(* IEC 61131-3 sources: Zbiorniki_user/Temp/Import/MpFile, 4 files *)

(* ---- MpFile.typ ---- *)
TYPE
	MpFileManagerUIItemType : 	STRUCT
		Name : STRING[255]; (*Filename / Folder name*)
		Size : UDINT; (*File size [bytes]*)
		LastModified : DATE_AND_TIME; (*Date when this file/folder was last modified*)
		ItemType : MpFileManagerUIItemTypeEnum; (*File type (.csv, .jpg, etc.)*)
		IsSelected : BOOL; (*Indicates that a file/folder is selected*)
		IsFolder : BOOL; (*Indicates that the element is a folder*)
	END_STRUCT;
	MpFileManagerUIItemTypeEnum :
		(
		mpFILE_ITEM_TYPE_NONE := 0, (*No type defined*)
		mpFILE_ITEM_TYPE_FOLDER := 1, (*Indicates that the element is a folder*)
		mpFILE_ITEM_TYPE_FILE := 2, (*Indicates that the element is a file*)
		mpFILE_ITEM_TYPE_TXT := 3, (*Indicates that the element is a text file*)
		mpFILE_ITEM_TYPE_HTML := 4, (*Indicates that the element is an HTML file*)
		mpFILE_ITEM_TYPE_DOC := 5, (*Indicates that the element is a Word file (.doc) *)
		mpFILE_ITEM_TYPE_XLS := 6, (*Indicates that the element is an Excel file (.xls)*)
		mpFILE_ITEM_TYPE_XML := 7, (*Indicates that the element is an XML file (.xml)*)
		mpFILE_ITEM_TYPE_CSV := 8, (*Indicates that the element is an CSV file (.csv)*)
		mpFILE_ITEM_TYPE_JPG := 9, (*Indicates that the element is an image file (.jpg)*)
		mpFILE_ITEM_TYPE_BMP := 10, (*Indicates that the element is an image file (.bmp)*)
		mpFILE_ITEM_TYPE_USER1 := 89, (*Indicates that the element is an user predefined type 1*)
		mpFILE_ITEM_TYPE_USER2 := 90, (*Indicates that the element is an user predefined type 2*)
		mpFILE_ITEM_TYPE_USER3 := 91, (*Indicates that the element is an user predefined type 3*)
		mpFILE_ITEM_TYPE_USER4 := 92, (*Indicates that the element is an user predefined type 4*)
		mpFILE_ITEM_TYPE_USER5 := 93, (*Indicates that the element is an user predefined type 5*)
		mpFILE_ITEM_TYPE_USER6 := 94, (*Indicates that the element is an user predefined type 6*)
		mpFILE_ITEM_TYPE_USER7 := 95, (*Indicates that the element is an user predefined type 7*)
		mpFILE_ITEM_TYPE_USER8 := 96, (*Indicates that the element is an user predefined type 8*)
		mpFILE_ITEM_TYPE_USER9 := 97, (*Indicates that the element is an user predefined type 9*)
		mpFILE_ITEM_TYPE_USER10 := 98, (*Indicates that the element is an user predefined type 10*)
		mpFILE_ITEM_TYPE_UNKNOWN := 99 (*Indicates that the file type is unknown*)
		);
	MpFileManagerUISortOrderEnum :
		(
		mpFILE_SORT_BY_NAME_ASC := 0, (*Sorts in ascending (alphabetic) order*)
		mpFILE_SORT_BY_NAME_DESC := 1, (*Sorts in descending (alphabetic) order*)
		mpFILE_SORT_BY_SIZE_ASC := 2, (*Sorts in ascending order by file size*)
		mpFILE_SORT_BY_SIZE_DES := 3, (*Sorts in descending order by file size*)
		mpFILE_SORT_BY_MOD_TIME_ASC := 4, (*Sorts in ascending order by date last modified*)
		mpFILE_SORT_BY_MOD_TIME_DESC := 5 (*Sorts in descending order by date last modified*)
		);
	MpFileManagerUIMessageEnum :
		(
		mpFILE_MSG_OK := 0, (*Dialog box for requesting confirmation of input*)
		mpFILE_MSG_CONFIRM_DELETE := 1, (*Dialog box for requesting confirmation of deletion*)
		mpFILE_MSG_CONFIRM_OVERWRITE := 2, (*Dialog box for requesting confirmation of overwriting*)
		mpFILE_MSG_BUSY := 3 (*Dialog box for requesting confirmation of busy UI*)
		);
	MpFileDiagType : 	STRUCT
		StatusID : MpFileStatusIDType; (*StatusID diagnostic structure*)
	END_STRUCT;
	MpFileStatusIDType : 	STRUCT
		ID : MpFileErrorEnum; (*Error code for mapp component*)
		Severity : MpComSeveritiesEnum; (*Describes the type of information supplied by the status ID (success, information, warning, error)*)
		Code : UINT; (*Code for the status ID. This error number can be used to search for additional information in the help system.*)
	END_STRUCT;
	MpFileInfoType : 	STRUCT
		Diag : MpFileDiagType; (*Diagnostic structure for the status ID*)
	END_STRUCT;
	MpFileManagerUIStatusEnum :
		(
		mpFILE_UI_STATUS_IDLE := 0, (*Indicates that no process is currently active*)
		mpFILE_UI_STATUS_REFRESH := 1, (*Updating elements*)
		mpFILE_UI_STATUS_CHANGE_PAGE := 2, (*Page change active*)
		mpFILE_UI_STATUS_CHANGE_DIR := 3, (*Folder change active*)
		mpFILE_UI_STATUS_CHANGE_DEVICE := 4, (*File Device Change active*)
		mpFILE_UI_STATUS_CREATE := 5, (*Creating a file/folder active*)
		mpFILE_UI_STATUS_RENAME := 6, (*Renaming a file/folder active*)
		mpFILE_UI_STATUS_DELETE := 7, (*Deleting a file/folder active*)
		mpFILE_UI_STATUS_COPY := 8, (*Copying a file/folder active*)
		mpFILE_UI_STATUS_CUT := 9, (*Cutting a file/folder active*)
		mpFILE_UI_STATUS_PASTE := 10, (*Pasting a file/folder active*)
		mpFILE_UI_STATUS_SORT := 11, (*Sorting files/folders in specified sort order*)
		mpFILE_UI_STATUS_ERROR := 99 (*The last operation generated an error*)
		);
	MpFileManagerUISetupType : 	STRUCT
		FileListSize : UINT := 10; (*Number of files to be displayed on one page of the list in the HMI application*)
		FileListScrollWindow : USINT := 1; (*Determines how many entries from the list are displayed in advance when scrolling up and down*)
	END_STRUCT;
	MpFileManagerUIConnectType : 	STRUCT
		Status : MpFileManagerUIStatusEnum; (*Current operation*)
		DeviceList : MpFileManagerUIDeviceListType; (*List of data storage media (file devices) accessible by the file manager*)
		File : MpFileManagerUIFileType; (*Contains the file list as well as additional information about files,folders and possible commands*)
		MessageBox : MpFileManagerUIMessageBoxType; (*Controls dialog boxes*)
		DefaultLayerStatus : UINT; (*Status DP for the default layer of the visu page where the file manager is being displayed*)
	END_STRUCT;
	MpFileManagerUIMessageBoxType : 	STRUCT
		LayerStatus : UINT; (*Visibility of the dialog box*)
		Type : MpFileManagerUIMessageEnum; (*Type of dialog box*)
		ErrorNumber : UINT; (*Current error number to be displayed*)
		Confirm : BOOL; (*Confirms the operation*)
		Cancel : BOOL; (*Cancels the operation*)
	END_STRUCT;
	MpFileManagerUIPathInfoType : 	STRUCT
		CurrentDir : STRING[255]; (*Current folder name*)
		FileCount : UDINT; (*Number of files in the current folder*)
		FolderCount : UDINT; (*Number of subfolders in the current folder*)
	END_STRUCT;
	MpFileManagerUIFileType : 	STRUCT
		List : MpFileManagerUIFileListType; (*List of all folders and files under the current path, as well as the navigation of the list*)
		Filter : STRING[255]; (*Filter used to sort the files*) (* *) (*#CMD#OPT#;*)
		SortOrder : MpFileManagerUISortOrderEnum; (*Responsible for the order of files in the list*)
		Refresh : BOOL; (*Updates the file list in the current folder*)
		PathInfo : MpFileManagerUIPathInfoType; (*Information about the current path*)
		EnterFolder : BOOL; (*Navigates one folder down*)
		FolderUp : BOOL; (*Navigates one folder up*)
		MultiSelect : BOOL; (*Allows the selection of multiple elements at the same time*)
		Delete : BOOL; (*Deletes a file or folder*)
		Copy : BOOL; (*Copying a file/folder*)
		Cut : BOOL; (*Cuts a file or folder*)
		Paste : BOOL; (*Pastes a file or folder*)
		NewName : STRING[255]; (*The new name of a file or folder when using the "Rename" or "CreateFolder" command*)
		Rename : BOOL; (*Renames a file or folder*)
		CreateFolder : BOOL; (*Creates a folder*)
	END_STRUCT;
	MpFileManagerUIFileListType : 	STRUCT
		Items : ARRAY[0..49]OF MpFileManagerUIItemType; (*List of all files and folders under the current path*)
		PageUp : BOOL; (*Jumps to the start of the current page and then scrolls up one page at a time*)
		StepUp : BOOL; (*Selects the previous entry in the list*)
		PageDown : BOOL; (*Jumps to the end of the current page and then scrolls down one page at a time*)
		StepDown : BOOL; (*Selects the next entry in the list*)
		RangeStart : REAL; (*Shows a bar indicating which part of the list is currently being displayed-Start [%]*)
		RangeEnd : REAL; (*Shows a bar indicating which part of the list is currently being displayed-End [%]*)
	END_STRUCT;
	MpFileManagerUIDeviceListType : 	STRUCT
		DeviceNames : ARRAY[0..9]OF STRING[50]; (*List of all available data storage media*)
		SelectedIndex : UINT; (*Index of the entry currently selected in the list*)
	END_STRUCT;
	MpFileManagerConfigType : 	STRUCT
		CustomizedFileType : ARRAY[0..9]OF STRING[5]; (*Customized file type names*)
	END_STRUCT;
END_TYPE

(* ---- MpFileAlarm.typ ---- *)
TYPE
	MpFileUIAlarmEnum :
		( (* Alarms of MpFile UI *)
		mpFILE_ALM_DEVICE_NOT_FOUND := 0, (*FileDevice not found*)
		mpFILE_ALM_ALREADY_EXISTING := 1, (*File/Folder already exists*)
		mpFILE_ALM_ERROR_FILE_SYSTEM := 2 (*General error in file system*)
		);
END_TYPE

(* ---- MpFileError.typ ---- *)
TYPE
    MpFileErrorEnum :
        ( (* Error numbers of library MpFile *)
        mpFILE_NO_ERROR := 0, (* No error *)
        mpFILE_ERR_ACTIVATION := -1064239103, (* Could not create component [Error: 1, 0xc0910001] *)
        mpFILE_ERR_MPLINK_NULL := -1064239102, (* MpLink is NULL pointer [Error: 2, 0xc0910002] *)
        mpFILE_ERR_MPLINK_INVALID := -1064239101, (* MpLink connection not allowed [Error: 3, 0xc0910003] *)
        mpFILE_ERR_MPLINK_CHANGED := -1064239100, (* MpLink modified [Error: 4, 0xc0910004] *)
        mpFILE_ERR_MPLINK_CORRUPT := -1064239099, (* Invalid MpLink contents [Error: 5, 0xc0910005] *)
        mpFILE_ERR_MPLINK_IN_USE := -1064239098, (* MpLink already in use [Error: 6, 0xc0910006] *)
        mpFILE_ERR_MISSING_UICONNECT := -1064165376, (* Missing value on UIConnect [Error: 8192, 0xc0922000] *)
        mpFILE_ERR_CMD_NOT_ALLOWED := -1064165375, (* Command {2:Command} not allowed [Error: 8193, 0xc0922001] *)
        mpFILE_ERR_NOTHING_TO_PASTE := -1064165374, (* No element to paste [Error: 8194, 0xc0922002] *)
        mpFILE_ERR_NOTHING_SELECTED := -1064165373, (* Nothing selected [Error: 8195, 0xc0922003] *)
        mpFILE_ERR_DIR_ALREADY_EXISTS := -1064165372, (* Folder {2:PathName} already exists in {3:DeviceName} [Error: 8196, 0xc0922004] *)
        mpFILE_ERR_INVALID_FILE_DEV := -1064165371, (* Invalid file device {2:DeviceName} [Error: 8197, 0xc0922005] *)
        mpFILE_ERR_NAME_EMPTY := -1064165370, (* New name not entered [Error: 8198, 0xc0922006] *)
        mpFILE_ERR_INVALID_NAME := -1064165369, (* Invaild name (ErrorCause: {1:ErrorNumber}) [Error: 8199, 0xc0922007] *)
        mpFILE_ERR_PASTE_NOT_ALLOWED := -1064165368, (* Paste not allowed (ErrorCause: {1:ErrorNumber}) [Error: 8200, 0xc0922008] *)
        mpFILE_ERR_FILE_SYSTEM := -1064165367, (* General error from file system (ErrorCause: {1:ErrorNumber}) [Error: 8201, 0xc0922009] *)
        mpFILE_ERR_INSUFF_ACCESS_RIGHT := -1064165358, (* User {2: UserName} has insufficient rights to access {3: Path} [Error: 8210, 0xc0922012] *)
        mpFILE_ERR_ITEM_IS_LOCKED := -1064165357, (* User {2: UserName} tried to access locked item {3: Path} (locked by user {4: LockUser}, since {5: LockTime}) [Error: 8211, 0xc0922013] *)
        mpFILE_ERR_COPY_ITEM := -1064165356, (* Item {3: SourcePath} could not be copied to {4: DestPath} (ErrorCause: {2: ErrorNumber}) [Error: 8212, 0xc0922014] *)
        mpFILE_ERR_ERASE_ITEM := -1064165355, (* Item {3: Path} could not be deleted (ErrorCause: {2: ErrorNumber}) [Error: 8213, 0xc0922015] *)
        mpFILE_ERR_INVALID_PATH := -1064165354, (* Invalid path-string {2: PathName} given [Error: 8214, 0xc0922016] *)
        mpFILE_ERR_INVALID_PARAMETER := -1064165353, (* Invalid parameter passed to function [Error: 8215, 0xc0922017] *)
        mpFILE_ERR_RENAME_ITEM := -1064165352, (* Item {3: Path} could not be renamed to {4: NewName} (ErorrCause: {2: ErrorNumber}) [Error: 8216, 0xc0922018] *)
        mpFILE_ERR_CREATE_ITEM := -1064165351, (* Item {3: Path} could not be created (ErrorCause: {2: ErrorNumber}) [Error: 8217, 0xc0922019] *)
        mpFILE_ERR_READ_ITEM := -1064165350, (* Item {3: Path} could not be read (ErrorCause: {2: ErrorNumber}) [Error: 8218, 0xc092201a] *)
        mpFILE_ERR_WRITE_ITEM := -1064165349, (* Item {3: Path} could not be written to (ErrorCause: {2: ErrorNumber}) [Error: 8219, 0xc092201b] *)
        mpFILE_INF_OVERWRITE := 1083318300 (* Item was overwritten [Informational: 8220, 0x4092201c] *)
        );
END_TYPE

(* ---- MpFile.fun ---- *)
FUNCTION_BLOCK MpFileManagerUI (*File management system and UI connection to VC4*) (* $GROUP=mapp Services,$CAT=File Explorer,$GROUPICON=Icon_mapp.png,$CATICON=Icon_MpFile.png *)
	VAR_INPUT
		MpLink : REFERENCE TO MpComIdentType; (*Connection to mapp*) (* *) (*#PAR#;*)
		Enable : BOOL; (*Enables/Disables the function block*) (* *) (*#PAR#;*)
		ErrorReset : BOOL; (*Resets function block errors*) (* *) (*#PAR#;*)
		UISetup : MpFileManagerUISetupType; (*Used to configure the elements connected to the HMI application*) (* *) (*#PAR#;*)
		UIConnect : REFERENCE TO MpFileManagerUIConnectType; (*This structure contains the parameters needed for the connection to the HMI application*) (* *) (*#CMD#;*)
	END_VAR
	VAR_OUTPUT
		Active : BOOL; (*Indicates whether the function block is active*) (* *) (*#PAR#;*)
		Error : BOOL; (*Indicates that the function block is in an error state or a command was not executed correctly*) (* *) (*#PAR#;*)
		StatusID : DINT; (*Status information about the function block*) (* *) (*#PAR#; *)
		Info : MpFileInfoType; (*Additional information about the component*) (* *) (*#CMD#;*)
	END_VAR
	VAR
		Internal : MpComInternalDataType; (*Internal stucture*)
	END_VAR
END_FUNCTION_BLOCK

FUNCTION_BLOCK MpFileManagerConfig (*mapp component for read/write component configuration*) (* $GROUP=mapp Services,$CAT=File Explorer,$GROUPICON=Icon_mapp.png,$CATICON=Icon_MpFile.png *)
	VAR_INPUT
		MpLink : REFERENCE TO MpComIdentType; (*Incoming communication handle (mapp standard interface)*) (* *) (*#PAR#;*)
		Enable : BOOL; (*Enables/Disables the function block (mapp standard interface)*) (* *) (*#PAR#;*)
		ErrorReset : BOOL; (*Resets all function block errors (mapp standard interface)*) (* *) (*#PAR#;*)
		Configuration : REFERENCE TO MpFileManagerConfigType; (*The component configuration structure.*) (* *) (*#PAR#; *)
		Load : BOOL; (*Reads the component configuration.*) (* *) (*#CMD#; *)
		Save : BOOL; (*Writes the component configuration.*) (* *) (*#CMD#; *)
	END_VAR
	VAR_OUTPUT
		Active : BOOL; (*Function block is active (mapp standard interface)*) (* *) (*#PAR#;*)
		Error : BOOL; (*Indicates an error (mapp standard interface)*) (* *) (*#PAR#;*)
		StatusID : DINT; (*Error/Status information (mapp standard interface)*) (* *) (*#PAR#; *)
		CommandBusy : BOOL; (*Function block is busy processing a command*) (* *) (*#CMD#OPT#;*)
		CommandDone : BOOL; (*True if a command finshed successfully.*) (* *) (*#CMD#;*)
		Info : MpFileInfoType; (*Provide any further useful information as function block output.(mapp standard interface)*) (* *) (*#CMD#; *)
	END_VAR
	VAR
		Internal : MpComInternalDataType; (*Internal data*)
	END_VAR
END_FUNCTION_BLOCK
